(* IEC 61131-3 sources: codesys-to-astra/src/POUs/F_C2aMbToReal, 2 files *)

(* ---- F_C2aMbToReal.decl.st ---- *)
// Назначение: два регистра Modbus (канал REGUL — ARRAY OF WORD, DPA-302.1 с. 15–16) -> REAL по порядку слов.
// Автор:      kr0nsch
// Версия:     0.1.0
// Документ:   docs/IO.md
FUNCTION F_C2aMbToReal : REAL
VAR_INPUT
    wFirst : WORD;              // первый регистр блока
    wSecond : WORD;             // второй регистр блока
    eOrder : E_C2aWordOrder;    // порядок слов
END_VAR
VAR
    uValue : U_C2aReal32;       // 32 бита как REAL/DWORD
END_VAR

(* ---- F_C2aMbToReal.impl.st ---- *)
IF eOrder = E_C2aWordOrder.LowWordFirst THEN
    uValue.dwValue := SHL(WORD_TO_DWORD(wSecond), 16) OR WORD_TO_DWORD(wFirst);  // lint:allow STL008 16 бит слова
ELSE
    uValue.dwValue := SHL(WORD_TO_DWORD(wFirst), 16) OR WORD_TO_DWORD(wSecond);  // lint:allow STL008 16 бит слова
END_IF
F_C2aMbToReal := uValue.rValue;
